(* PLC project TBEN_L5_PLC11.project, CODESYS CODESYS V3.5 SP21 Patch 1 *)
(* stored: creationDateTime 2026-11-07T15:34:50.2258646, modificationDateTime 2026-11-07T15:09:07.4034196 *)

{attribute 'qualified_only'}
// Giá trị byte Control của khung IOL_CALL (request)
TYPE E_IolService :
(
    WRITE := 2,   // ISDU write
    READ  := 3    // ISDU read
) USINT;
END_TYPE
